Fanuc KAREL source: kd00015.KL

-- PROVISIONAL review KL for V1013-1; original PC SHA256 c4bef491dfea5bb1d98affd5a0cf610db081f7e2987b4ae7926769c924b3e875
-- Incomplete behavior may be omitted. Consult companion uncertainty JSON. Do not deploy.
PROGRAM KD00015
%NOLOCKGROUP
VAR
  I : INTEGER
  J : INTEGER
  B : BOOLEAN
  R : REAL
  S : STRING[80]
BEGIN
  -- UNRESOLVED_PC offsets 5-6; opcodes 16
  -- UNRESOLVED_PC offsets 11-15; opcodes 7F
END KD00015
